Staubli VAL3: onSave.pgx

public program onSave(bool& x_bTosave)
begin
  if x_bTosave
    rs:bIsSaving=true
    progTemp:libSave()
    x_bTosave=false
    rs:bIsSaving=false
    delay(0.1)
    popUpMsg("数据已保存")
  endIf
end
